(* IEC 61131-3 sources: JingjiangMoonbox/Application/Application/任务列表/Main_Task/GNS_MAP/STRUCT, 2 files *)

(* ---- StSysGantryAxisInf.st ---- *)
(*@CES
Name=StSysGantryAxisInf
Type=Gvl
TypeGuid=2db5746d-d284-4425-9f7f-2663a34b0ebc
Guid=7a9ba2fe-c896-4159-a4c9-1568d21622d8
HasDeclaration=True
HasImplementation=False
*)
{DECLARATION}
TYPE StSysGantryAxisInf :(*系统龙门轴信息@总共20个龙门轴*)
STRUCT
	byGantryAxisNum:BYTE;(*龙门轴总数*)
	astGantryAxisInf:ARRAY [1..20] OF StGantryAxisInf;
END_STRUCT
END_TYPE
{IMPLEMENTATION}

(* ---- StSysStationInf.st ---- *)
(*@CES
Name=StSysStationInf
Type=Gvl
TypeGuid=2db5746d-d284-4425-9f7f-2663a34b0ebc
Guid=ff62fd15-378a-4887-af92-0b6cfd3f9fba
HasDeclaration=True
HasImplementation=False
*)
{DECLARATION}
TYPE StSysStationInf :(*系统的站信息@最大128个站*)
STRUCT
	byStationNum:BYTE;
	astStationInf:ARRAY [1..128] OF StStationInf;
END_STRUCT
END_TYPE

{IMPLEMENTATION}
